{attribute 'qualified_only'}
{attribute 'to_string'}
TYPE E_AutomaticExtractionState :
(
	AUTO_EXTRACTION := 0,
	REDUCE_PUMP_START_CALIB := 1,
	WAIT_FOR_PRESSURE_REDUCE := 2,
	CLOSE_ON_OFF_VALVE := 3,
	FILLING_ACTIVE := 4,
	WAIT_FOR_PRESSURE_TO_SET := 5,
	INCREASE_PUMP := 6,
	OPEN_ON_OFF_VALVE := 7,
	MANUAL_EXTRACTION := 8
	
);
END_TYPE

(* stored: Version 1.1.0.1, ProductVersion 3.1.4024.9
   DUT E_AutomaticExtractionState: Id {4f6d5abb-7cc1-48dc-88f2-3a80d66f4e1e} *)
